// TIA Portal V21 export
// export: Created 2026-11-21T13:26:58.9491956Z, ExportSetting WithDefaults, DisplayName Totally Integrated Automation Portal, DisplayVersion V21, DisplayName STEP 7 Professional, DisplayVersion V21, DisplayName STEP 7 Safety, DisplayVersion V21, DisplayName Tech WebApplication, DisplayVersion V21, DisplayName WinCC Basic/Comfort/Advanced, DisplayVersion V21, DisplayName WinCC Unified, DisplayVersion V21
DATA_BLOCK "Recipe"   // DB30
TITLE = Rezept / Recipe / Recette
{ S7_Optimized_Access := 'TRUE' }
VERSION : 0.1
// Werte des Rezepts / Values of the recipe / Valeurs de la recette
// stored: AutoNumber true, DBAccessibleFromOPCUA true, DBAccessibleFromWebserver true, IsOnlyStoredInLoadMemory false, IsRetainMemResEnabled false, IsWriteProtectedInAS false, MemoryReserve 100
   VAR
      target : Int := 500;   // Sollfüllstand in mm / Target level in mm / Niveau de consigne en mm
      hysteresis : Int := 20;   // Hysteresis in mm
   END_VAR
BEGIN
END_DATA_BLOCK
